(* IEC 61131-3 sources: SemaPLC/sema-plc-benchmark/spec2control-benchmark/data/st-baseline/multi-phase-flow-facility/pous/programs, 7 files *)

(* ---- main.st ---- *)
PROGRAM main
VAR
	Heartbeat : bool;
END_VAR

(* Entry point required by OpenPLC Editor v4. The process sections run as parallel program instances under task0; main only provides a scan heartbeat. *)
Heartbeat := NOT Heartbeat;

END_PROGRAM

(* ---- Section2.st ---- *)
PROGRAM Section2
VAR
	FT404_GasFlow_PV : real;
	FT406_LiqFlow_PV : real;
	PT403_SepPressure_PV : real;
	PT408_AuxPressure_PV : real;
	FIC406_LiqFlow_SP_From_FFIC402 : real;
	FT_404 : ANALOG_IN;
	FT_406 : ANALOG_IN;
	PT_403 : ANALOG_IN;
	PT_408 : ANALOG_IN;
	FFIC_402 : RATIO_CONTROL;
	FIC_406 : PID_BASIC;
	PIC_401 : PID_BASIC;
	CV_406 : VALVE_ELECTRIC;
	CV_401 : VALVE_ELECTRIC;
	ValveInhibit_OR : bool;
	RatioInhibit_OR : bool;
END_VAR

FT_404(
    PV_Low := 50.0);
FT_406(
    PV_Low := 20.0);
PT_403();
PT_408();
RatioInhibit_OR := PT_403.High_Alarm OR PT_403.Low_Alarm OR FT_404.Low_Alarm OR FT_404.General_Fault OR FT_406.General_Fault OR PT_408.Low_Alarm;
FFIC_402(
    Auto := TRUE,
    PrimaryPV := FT_404.PV,
    SecondaryPV := FT_406.PV,
    RatioSP := 2.5,
    MV_MIN := 0.0,
    MV_MAX := 500.0,
    Inhibit := RatioInhibit_OR);
FIC_406(
    AUTO := TRUE,
    PV := FT_406.PV,
    SP := FFIC_402.SlaveSP);
PIC_401(
    AUTO := TRUE,
    PV := PT_403.PV,
    SP := 5.0,
    PV_High := 6.0,
    PV_Low := 4.0);
ValveInhibit_OR := PT_403.High_Alarm OR PT_403.Low_Alarm OR FT_404.Low_Alarm OR FT_406.Low_Alarm;
CV_406(
    Control_Signal := FIC_406.XOUT,
    Inhibit := ValveInhibit_OR);
CV_401(
    Control_Signal := PIC_401.XOUT);

(* Outputs published to other sections / HMI. *)
FT404_GasFlow_PV := FT_404.PV;
FT406_LiqFlow_PV := FT_406.PV;
PT403_SepPressure_PV := PT_403.PV;
PT408_AuxPressure_PV := PT_408.PV;
FIC406_LiqFlow_SP_From_FFIC402 := FFIC_402.SlaveSP;

END_PROGRAM

(* ---- Section3.st ---- *)
PROGRAM Section3
VAR
	PT501_Pressure_PV : real;
	LI502_Level_PV : real;
	PIC501_Output_To_FV102 : real;
	PT_501 : ANALOG_IN;
	LI_502 : ANALOG_IN;
	PIC_501 : PID_BASIC;
	FV_102 : VALVE_ELECTRIC;
	SeparatorShutdown_OR : bool;
	PIC501_Inhibit_OR : bool;
END_VAR

PT_501(
    PV_High := 85.0,
    PV_Low := 65.0,
    Scaling_Slope := 9.375,
    Scaling_Offset := -37.5);
LI_502(
    PV_High := 90.0,
    PV_Low := 5.0,
    Scaling_Slope := 6.25,
    Scaling_Offset := -25.0);
SeparatorShutdown_OR := PT_501.General_Fault OR PIC_501.PV_High_Alarm;
FV_102(
    Control_Signal := PIC_501.XOUT,
    Manual_Mode := FALSE,
    Open_Limit := 100.0,
    Close_Limit := 0.0,
    Inhibit := SeparatorShutdown_OR);
PIC501_Inhibit_OR := SeparatorShutdown_OR OR PT_501.High_Alarm OR PT_501.Low_Alarm OR LI_502.Low_Alarm OR LI_502.High_Alarm OR FV_102.Alarm;
PIC_501(
    AUTO := TRUE,
    PV := PT_501.PV,
    SP := 75.0,
    MV_MIN := 0.0,
    MV_MAX := 100.0,
    X0 := FV_102.Feedback_Pos,
    KP := 2.0,
    TR := 0.5,
    TD := 0.1,
    Inhibit := PIC501_Inhibit_OR);

(* Outputs published to other sections / HMI. *)
PT501_Pressure_PV := PT_501.PV;
LI502_Level_PV := LI_502.PV;
PIC501_Output_To_FV102 := PIC_501.XOUT;

END_PROGRAM

(* ---- Section4.st ---- *)
PROGRAM Section4
VAR
	LI201_Raw_mA : real;
	XV010_OpenSw_Raw : bool;
	XV011_OpenSw_Raw : bool;
	LI201_Level_PV_Pct : real;
	FIC302_MV_To_FV101_Pct : real;
	FV101_Feedback_Position_Pct : real;
	FIC_302 : PID_BASIC;
	FV_101 : VALVE_ELECTRIC;
	LI_201 : ANALOG_IN;
	XV_010_OPEN_FB : DIGITAL_IN;
	XV_011_OPEN_FB : DIGITAL_IN;
	FlowPathOpen_AND : bool;
	NotFlowPathOpen_NOT : bool;
	FV101ManualMode_OR : bool;
	LIFaultInvert_NOT : bool;
	LoopAutoPermissive_AND : bool;
END_VAR

LI_201(
    Raw_Signal := LI201_Raw_mA,
    PV_High := 80.0,
    PV_Low := 20.0,
    Scaling_Slope := 6.25,
    Scaling_Offset := -25.0);
XV_010_OPEN_FB(
    DI_Raw := XV010_OpenSw_Raw);
XV_011_OPEN_FB(
    DI_Raw := XV011_OpenSw_Raw);
FlowPathOpen_AND := XV_010_OPEN_FB.DI_Out AND XV_011_OPEN_FB.DI_Out;
LIFaultInvert_NOT := NOT LI_201.General_Fault;
LoopAutoPermissive_AND := LIFaultInvert_NOT AND FlowPathOpen_AND;
FIC_302(
    AUTO := LoopAutoPermissive_AND,
    PV := LI_201.PV,
    SP := 70.0,
    MV_MIN := 0.0,
    MV_MAX := 100.0,
    X0 := 25.0,
    KP := 1.8,
    TR := 2.0,
    TD := 0.3);
NotFlowPathOpen_NOT := NOT FlowPathOpen_AND;
FV101ManualMode_OR := NotFlowPathOpen_NOT OR FIC_302.PV_High_Alarm;
FV_101(
    Control_Signal := FIC_302.XOUT,
    Manual_Mode := FV101ManualMode_OR,
    Manual_Position := 0.0,
    Open_Limit := 100.0,
    Close_Limit := 0.0);

(* Outputs published to other sections / HMI. *)
LI201_Level_PV_Pct := LI_201.PV;
FIC302_MV_To_FV101_Pct := FIC_302.XOUT;
FV101_Feedback_Position_Pct := FV_101.Feedback_Pos;

END_PROGRAM

(* ---- Section5.st ---- *)
PROGRAM Section5
VAR
	FIC101_MV_PCT : real;
	FIC102_MV_PCT : real;
	P001_Speed_AO_PCT : real;
	P001_Start_Cmd : bool;
	P001_Stop_Cmd : bool;
	FT102_FlowOK_Thresh : real;
	ValveOpenFB_Threshold : real;
	LevelOK_Threshold : real;
	FIC101_Deviation_Alarm_15s : bool;
	FIC102_Deviation_Alarm_15s : bool;
	FT_102 : ANALOG_IN;
	FT_104 : ANALOG_IN;
	LI_101 : ANALOG_IN;
	FIC_101 : PID_BASIC;
	FIC_102 : PID_BASIC;
	FV_103 : VALVE_ELECTRIC;
	P_001 : MOTOR_VSD;
	FlowOK_TON : TON;
	FIC101_Dev_TON : TON;
	FIC102_Dev_TON : TON;
	FIC101_ForceManual_OR : bool;
	FIC102_ForceManual_OR : bool;
	FIC101_AutoEnable_NOT : bool;
	FIC102_AutoEnable_NOT : bool;
	FT102_GT_10GPM : bool;
	ValveOpenPermissive_AND : bool;
	ValveOpenInhibit_NOT : bool;
	ValveInhibit_OR : bool;
	LevelOK_GT25 : bool;
	ValveFB_GT_90PCT : bool;
	P001_StartPermissive_AND : bool;
	P001_Stop_OR : bool;
END_VAR

(* Constant configuration values. *)
FT102_FlowOK_Thresh := 10.0;
ValveOpenFB_Threshold := 90.0;
LevelOK_Threshold := 25.0;

FT_102(
    Scaling_Slope := 6.25,
    Scaling_Offset := -25.0);
FT_104(
    Scaling_Slope := 6.25,
    Scaling_Offset := -25.0);
LI_101(
    PV_High := 90.0,
    PV_Low := 20.0,
    Scaling_Slope := 6.25,
    Scaling_Offset := -25.0);
FIC101_ForceManual_OR := LI_101.Low_Alarm OR LI_101.High_Alarm OR FT_102.General_Fault;
FIC101_AutoEnable_NOT := NOT FIC101_ForceManual_OR;
FIC_101(
    AUTO := FIC101_AutoEnable_NOT,
    PV := FT_102.PV,
    SP := 50.0,
    MV_MIN := 0.0,
    MV_MAX := 100.0,
    X0 := 0.0,
    KP := 2.0,
    TR := 1.0,
    TD := 0.1,
    Deviation_Limit := 10.0);
FIC102_ForceManual_OR := LI_101.Low_Alarm OR LI_101.High_Alarm OR FT_104.General_Fault;
FIC102_AutoEnable_NOT := NOT FIC102_ForceManual_OR;
FIC_102(
    AUTO := FIC102_AutoEnable_NOT,
    PV := FT_104.PV,
    SP := 45.0,
    MV_MIN := 0.0,
    MV_MAX := 100.0,
    X0 := 0.0,
    KP := 2.0,
    TR := 1.0,
    TD := 0.1,
    Deviation_Limit := 8.0);
FT102_GT_10GPM := (FT_102.PV > FT102_FlowOK_Thresh);
FlowOK_TON(
    IN := FT102_GT_10GPM,
    PT := T#8s);
LevelOK_GT25 := (LI_101.PV > LevelOK_Threshold);
ValveFB_GT_90PCT := (FV_103.Feedback_Pos > ValveOpenFB_Threshold);
P001_StartPermissive_AND := P001_Start_Cmd AND LevelOK_GT25 AND ValveFB_GT_90PCT;
P001_Stop_OR := P001_Stop_Cmd OR LI_101.General_Fault;
P_001(
    Start_Cmd := P001_StartPermissive_AND,
    Stop_Cmd := P001_Stop_OR,
    Speed_SP := FIC_102.XOUT,
    Inhibit := LI_101.General_Fault);
ValveOpenPermissive_AND := P_001.FB_Running AND FlowOK_TON.Q;
ValveOpenInhibit_NOT := NOT ValveOpenPermissive_AND;
ValveInhibit_OR := ValveOpenInhibit_NOT OR LI_101.General_Fault;
FV_103(
    Control_Signal := FIC_101.XOUT,
    Manual_Mode := FALSE,
    Manual_Position := 0.0,
    Open_Limit := 25.0,
    Close_Limit := 0.0,
    Inhibit := ValveInhibit_OR);
FIC101_Dev_TON(
    IN := FIC_101.Deviation_Alarm,
    PT := T#15s);
FIC102_Dev_TON(
    IN := FIC_102.Deviation_Alarm,
    PT := T#15s);

(* Outputs published to other sections / HMI. *)
FIC101_Deviation_Alarm_15s := FIC101_Dev_TON.Q;
FIC102_Deviation_Alarm_15s := FIC102_Dev_TON.Q;
FIC101_MV_PCT := FIC_101.XOUT;
FIC102_MV_PCT := FIC_102.XOUT;
P001_Speed_AO_PCT := P_001.Speed_Out;

END_PROGRAM

(* ---- Section6.st ---- *)
PROGRAM Section6
VAR
	FT105_FlowRate_gpm : real;
	LI503_Level_Pct : real;
	P001_Running_Permissive : bool;
	FT_105 : ANALOG_IN;
	LI_503 : ANALOG_IN;
	LIC_502 : PID_BASIC;
	LIC_503 : PID_BASIC;
	LVC_502 : VALVE_ELECTRIC;
	LVC_507 : VALVE_ELECTRIC;
	P_001 : MOTOR_ON_OFF;
	PumpNotRunning : bool;
	LevelOverride : bool;
	FlowOverride : bool;
END_VAR

FT_105(
    PV_High := 45.0,
    PV_Low := 5.0,
    Scaling_Slope := 3.125,
    Scaling_Offset := -12.5,
    Alarm_Enable := TRUE);
LI_503(
    PV_High := 90.0,
    PV_Low := 10.0,
    Scaling_Slope := 6.25,
    Scaling_Offset := -25.0,
    Alarm_Enable := TRUE);
P_001();
PumpNotRunning := NOT P_001.FB_Running;
FlowOverride := FT_105.Low_Alarm OR FT_105.High_Alarm OR PumpNotRunning OR FT_105.General_Fault;
LIC_502(
    AUTO := TRUE,
    PV := FT_105.PV,
    SP := 35.0,
    MV_MIN := 0.0,
    MV_MAX := 100.0,
    KP := 1.8,
    TR := 2.0,
    TD := 0.0,
    Inhibit := FlowOverride);
LevelOverride := LI_503.High_Alarm OR LI_503.Low_Alarm OR PumpNotRunning OR LI_503.General_Fault;
LIC_503(
    AUTO := TRUE,
    PV := LI_503.PV,
    SP := 65.0,
    MV_MIN := 0.0,
    MV_MAX := 100.0,
    KP := -2.0,
    TR := 1.5,
    TD := 0.1,
    Inhibit := LevelOverride);
LVC_502(
    Control_Signal := LIC_502.XOUT,
    Manual_Mode := FlowOverride,
    Manual_Position := 100.0,
    Open_Limit := 100.0,
    Close_Limit := 0.0,
    Inhibit := FlowOverride);
LVC_507(
    Control_Signal := LIC_503.XOUT,
    Manual_Mode := LevelOverride,
    Manual_Position := 0.0,
    Open_Limit := 100.0,
    Close_Limit := 0.0,
    Inhibit := LevelOverride);

(* Outputs published to other sections / HMI. *)
FT105_FlowRate_gpm := FT_105.PV;
LI503_Level_Pct := LI_503.PV;
P001_Running_Permissive := P_001.FB_Running;

END_PROGRAM

(* ---- Section7.st ---- *)
PROGRAM Section7
VAR
	PIT106_Raw_mA : real;
	CompressorRunPermissive : bool;
	PIT106_PressureBar : real;
	PIC105_MV_Percent : real;
	PIT_106 : ANALOG_IN;
	COMP_RUN_PERM : BOOL_INPUT;
	PIC_105 : PID_BASIC;
	V_010 : VALVE_ELECTRIC;
	CompStartupDelay : TON;
	CompNotRunning : bool;
	AirCompInhibit : bool;
	StartupNotElapsed : bool;
END_VAR

PIT_106(
    Raw_Signal := PIT106_Raw_mA,
    PV_High := 9.5,
    PV_Low := 0.5,
    Scaling_Slope := 0.625,
    Scaling_Offset := -2.5);
COMP_RUN_PERM(
    Bool_In := CompressorRunPermissive);
CompNotRunning := NOT COMP_RUN_PERM.Bool_Out;
CompStartupDelay(
    IN := COMP_RUN_PERM.Bool_Out,
    PT := T#7s);
StartupNotElapsed := NOT CompStartupDelay.Q;
AirCompInhibit := CompNotRunning OR PIT_106.High_Alarm OR PIT_106.Low_Alarm OR PIT_106.General_Fault OR StartupNotElapsed;
PIC_105(
    AUTO := TRUE,
    PV := PIT_106.PV,
    SP := 8.5,
    MV_MIN := 0.0,
    MV_MAX := 100.0,
    KP := 3.0,
    TR := 1.2,
    TD := 0.3,
    Inhibit := AirCompInhibit);
V_010(
    Control_Signal := PIC_105.XOUT,
    Manual_Mode := FALSE,
    Open_Limit := 100.0,
    Close_Limit := 0.0,
    Inhibit := AirCompInhibit);

(* Outputs published to other sections / HMI. *)
PIT106_PressureBar := PIT_106.PV;
PIC105_MV_Percent := PIC_105.XOUT;

END_PROGRAM
